Fanuc KAREL source: kt00165.KL

-- PROVISIONAL review KL for V770-1; original PC SHA256 a115d8dcaa75b0858f8d3cf3b37524568ef9fa483dc23f7ee831995e446ff9d4
-- Incomplete behavior may be omitted. Consult companion uncertainty JSON. Do not deploy.
PROGRAM KT00165
%NOLOCKGROUP
VAR
  I1 : INTEGER
  OUT : INTEGER
-- UNRESOLVED_DECL Y2 type=002018
BEGIN
  -- UNRESOLVED_PC offsets 5-16; opcodes 2E,23
  -- UNRESOLVED_PC offsets 21-35; opcodes 2E,22,9D,33,B2
  -- UNRESOLVED_PC offsets 40-62; opcodes 21,22,9D,33,B1,56,23
  -- UNRESOLVED_PC offsets 67-71; opcodes 7F
END KT00165
